(* IEC 61131-3 sources: Piper/src/Ar/MachineControl/MachineProg, 5 files *)

(* ---- MachineProg.typ ---- *)
(*
* File: MachineProg.typ
* Copyright (c) 2023 Loupe
* https://loupe.team
*
* This file is part of MachineProg, licensed under the MIT License.
*)

TYPE
	Configuration_typ : 	STRUCT
		remotePLC : BOOL;
	END_STRUCT;
END_TYPE

(* ---- ApplicationCodeExample.st ---- *)
// In this example, the network used is powerlink, and there is one main with one remote.

ACTION CommsVerifySize:

	// Verify the size of IO variables used in multi-PLC communication.

	SIZEOF_MODULE_MAIN := SIZEOF(gMachine.IO.oMainInterface);
	SIZEOF_MODULE_REMOTE := SIZEOF(gMachine.IO.iMainInterface);

	IF SIZEOF(gMachine.IO.oMainInterface) = SIZEOF(oModuleInterface)
		AND SIZEOF(gMachine.IO.iMainInterface) = SIZEOF(iModuleInterface) THEN
		ioSizeVerfied := TRUE;
	ELSE
		logError('App', 0, 'Piper IO interface does not match buffer size. Comms disabled.', 0);
		//errcolAddError(ADR('MachineProg'), ADR('Piper IO interface does not match buffer size. Comms disabled.'), 0, 0, gErrorCollector);
	END_IF

END_ACTION

ACTION CommsHandleInputs:

	// Write the input IO to the appropriate module interface

	IF ioSizeVerfied AND iNetworkConnected THEN
		IF Configuration.remotePLC THEN
			brsmemcpy(ADR(gMachine.IO.iMainInterface), ADR(iModuleInterface), SIZEOF_MODULE_REMOTE);
		ELSE
			brsmemcpy(ADR(remoteModuleInterface), ADR(iModuleInterface), SIZEOF_MODULE_REMOTE);
		END_IF
	END_IF

END_ACTION

ACTION CommsHandleOutputs:

	// Write the appropriate module interface to the output IO

	IF ioSizeVerfied THEN
		IF Configuration.remotePLC THEN
			brsmemcpy(ADR(oModuleInterface), ADR(gMachine.IO.oMainInterface), SIZEOF_MODULE_MAIN);
		ELSE
			brsmemcpy(ADR(oModuleInterface), ADR(remoteModuleInterface), SIZEOF_MODULE_MAIN);
		END_IF
	END_IF

END_ACTION

ACTION CommsHandleNetwork:

	// Handle network connects and disconnects

	powerLinkConnectedRTrig.CLK := iNetworkConnected;
	powerLinkConnectedRTrig();

	powerLinkConnectedFTrig.CLK := iNetworkConnected;
	powerLinkConnectedFTrig();

	IF remoteModuleErrorAck THEN
		remoteModuleErrorAck := FALSE;
		remoteModuleError := FALSE;
	END_IF

	IF ioSizeVerfied THEN
		IF Configuration.remotePLC THEN
			IF NOT gIsRemote THEN
				IF NOT gMachine.IO.iMainInterface.ModuleIsBypassed THEN
					gIsRemote := TRUE;
				END_IF
			END_IF

			// TODO: Handle powerlink disconnects better
			IF powerLinkConnectedFTrig.Q THEN // TODO: Do we need a debounce for this?
				// IF we loose connection while running, stop
				gIsRemote := FALSE;
				gMachine.IN.CMD.Abort := TRUE;
			END_IF

			remoteModuleInterface.ModuleBypass := TRUE; // We want to ingore our selves with we are changed to a remote :)
		ELSE

			IF remoteModuleInterface.ModuleName = '' THEN
				remoteModuleInterface.ModuleName := 'Remote PLC';
			END_IF

			IF powerLinkConnectedFTrig.Q THEN
				IF NOT remoteModuleInterface.ModuleBypass THEN
					IF gMachine.OUT.State <> MACH_ST_ABORTED THEN
						gMachine.IN.CMD.Abort := TRUE;
					END_IF

				END_IF
				// TODO: We will need to handle reconnects
				remoteModuleInterface.ModuleBypass := TRUE; // Disconnect remote from Piper
			END_IF

			IF remoteModuleInterface.ModuleBypass THEN
				// TODO: gMachine.IO.oModule is not populated while acting as a main Piper, so remoteModuleInterface.PiperState will not be updated while bypassed. So This will not work until we fix that
				IF iNetworkConnected AND gMachine.OUT.State = MACH_ST_ABORTED AND remoteModuleInterface.PiperState = MACH_ST_ABORTED THEN // remoteModuleInterface only represents the remote until piper is called
					remoteModuleInterface.ModuleBypass := FALSE; // Connect remote to Piper
				END_IF

				IF NOT remoteModuleError THEN
					remoteModuleError := TRUE; // Error latch so we dont spam errors
					logError('App', 0, 'Module disconnected from powerlink', 0);
					//errcolAddError(ADR(remoteModuleInterface.ModuleName), ADR('Module disconnected from powerlink'), 0, ADR(remoteModuleErrorAck), gErrorCollector);
				END_IF
			END_IF

			remoteModule.ModuleInterface := ADR(remoteModuleInterface);
			remoteModule.Piper := ADR(gMachine);
			remoteModule();

			// Temp fix because Piper remote does not handle boot right now
			IF gMachine.OUT.State = MACH_ST_BOOTING THEN
				remoteModuleInterface.ModuleResponse := MACH_ST_BOOTING;
			END_IF
		END_IF
	END_IF

END_ACTION

(* ---- ApplicationCodeExample.var ---- *)
(********************************************************************
 * COPYRIGHT -- Automation Resources Group
 ********************************************************************
 * Program: MachineProg
 * File: MachineProg.var
 * Author: David Blackburn
 * Created: November 10, 2011
 ********************************************************************
 * Local variables of program MachineProg
 ********************************************************************)
VAR
	powerLinkConnectedRTrig : R_TRIG;
	powerLinkConnectedFTrig : F_TRIG;
	iNetworkConnected : BOOL;
	remoteModule : Piper_Module_Fub;
	remoteModuleInterface : Module_Interface_typ;
	SIZEOF_MODULE_MAIN : UDINT;
	SIZEOF_MODULE_REMOTE : UDINT;
	ioSizeVerfied : BOOL;
	iModuleInterface : ARRAY[0..195] OF USINT;
	oModuleInterface : ARRAY[0..195] OF USINT;
	remoteModuleErrorAck : BOOL;
	remoteModuleError : BOOL;
END_VAR

(* ---- MachineProgCyclic.st ---- *)
(*
* File: MachineProgCyclic.st
* Copyright (c) 2023 Loupe
* https://loupe.team
*
* This file is part of MachineProg, licensed under the MIT License.
*)

PROGRAM _INIT

	gIsRemote := Configuration.remotePLC;

	CommsVerifySize;

END_PROGRAM

PROGRAM _CYCLIC

	CommsHandleInputs;

	CommsHandleNetwork; // This needs to be after CommsHandleInputs, but before Piper is called

	//Piper controls the main machine state
	Piper_Remote_fn_Cyclic( gMachine, gIsRemote );

	//Handle anything that needs to happen at the machine level for a given state
	CASE gMachine.OUT.State OF

		MACH_ST_BOOTING:
			StateString:= 'Booting';
			TON_0.IN:=	1;

		MACH_ST_BOOTED:
			StateString:= 'Booted';
			IF TON_0.IN THEN
				TON_0.IN:=	0;
				IF BootTime = 0 THEN
					BootTime:= TON_0.ET;
				END_IF
				BootTime:= 	(TON_0.ET+(BootTime*9))/10;
			END_IF
		MACH_ST_NOT_READY :StateString:= 'MACH_ST_NOT_READY';
		MACH_ST_ERROR	  :StateString:= 'MACH_ST_ERROR	;  ';
		MACH_ST_CLEARING  :StateString:= 'MACH_ST_CLEARING ';
		MACH_ST_STOPPED	  :StateString:= 'MACH_ST_STOPPED  ';
		MACH_ST_STARTING  :StateString:= 'MACH_ST_STARTING ';
		MACH_ST_IDLE	  :StateString:= 'MACH_ST_IDLE     ';
		MACH_ST_SUSPENDED :StateString:= 'MACH_ST_SUSPENDED';
		MACH_ST_EXECUTE	  :StateString:= 'MACH_ST_EXECUTE  ';
		MACH_ST_STOPPING  :StateString:= 'MACH_ST_STOPPING ';
		MACH_ST_ABORTING  :StateString:= 'MACH_ST_ABORTING ';
		MACH_ST_ABORTED	  :StateString:= 'MACH_ST_ABORTED  ';
		MACH_ST_HOLDING	  :StateString:= 'MACH_ST_HOLDING  ';
		MACH_ST_HELD	  :StateString:= 'MACH_ST_HELD     ';
		MACH_ST_UNHOLDING :StateString:= 'MACH_ST_UNHOLDING';
		MACH_ST_SUSPENDING:StateString:= 'MACH_ST_SUSPENDING';
		MACH_ST_UNSUSPENDING:StateString:= 'MACH_ST_UNSUSPENDING';
		MACH_ST_RESETTING :StateString:= 'MACH_ST_RESETTING';
		MACH_ST_COMPLETING:StateString:= 'MACH_ST_COMPLETING';
		MACH_ST_COMPLETE  :StateString:= 'MACH_ST_COMPLETE ';
		MACH_ST_BYPASSED  :StateString:= 'MACH_ST_BYPASSED ';
		MACH_ST_		  :StateString:= 'MACH_ST_	       ';
	END_CASE

	CASE gMachine.OUT.State OF
		MACH_ST_STARTING,
		MACH_ST_EXECUTE,
		MACH_ST_HELD,
		MACH_ST_UNHOLDING,
		MACH_ST_SUSPENDING,
		MACH_ST_UNSUSPENDING,
		MACH_ST_HOLDING,
		MACH_ST_COMPLETING,
		MACH_ST_COMPLETE:
			//Mode change not allowed
			gRequestedMode:=gActiveMode;
		ELSE
			gActiveMode:=gRequestedMode;
	END_CASE

	TON_0.PT:=T#1d;
	TON_0();

	//**************************************************************************//
	//Display the first module the Piper is waiting on							//
	//**************************************************************************//
	IF gMachine.OUT.BusyModule = 0 THEN
		StatusModule.ModuleName:=	'Ready';
		Module ACCESS ADR(StatusModule);
	ELSE
		Module ACCESS gMachine.OUT.BusyModule;
		StatusModule:= Module;
	END_IF;

	CommsHandleOutputs;

END_PROGRAM

(* ---- MachineProg.var ---- *)
(*
* File: MachineProg.var
* Copyright (c) 2023 Loupe
* https://loupe.team
*
* This file is part of MachineProg, licensed under the MIT License.
*)

VAR
	StatusModule : Module_Interface_typ;
	Module : REFERENCE TO Module_Interface_typ;
	TON_0 : TON;
	StateString : STRING[80];
END_VAR
VAR RETAIN
	ByPassAll : BOOL := 0;
END_VAR
VAR
	Configuration : Configuration_typ;
END_VAR
